// TIA Portal V18 export
DATA_BLOCK "MCP_RC_DB3"   // DB9803
{ S7_Optimized_Access := 'TRUE' }
   VAR
      Count : Int := 5;
      Grp : Struct
         Inner : "MCP_RC_UDT";
         Flag : Bool := TRUE;
      END_STRUCT;
   END_VAR
BEGIN
   Grp.Inner.Speed := 12;
END_DATA_BLOCK
